(* IEC 61131-3 sources: brOscatLib/oscatBasic (part 4) *)

(* ---- FADE.st ---- *)
FUNCTION_BLOCK FADE
    (*http://www.oscat.de/images/OSCATBasic/oscat_basic333_en.pdf#page=276*)
    rmx(RST := RST AND NOT F, SET := RST AND F, PT := TF, UP := F);
    Y := (IN2 - IN1) / 65535.0 * WORD_TO_REAL(rmx.OUT) + IN1;

    (* code for rev 1.1
    IF RST THEN
    	rmx(set := F, RST := NOT F);
    ELSIF F AND (NOT rmx.high) THEN
    	rmx(PT := TF, UP := TRUE, e := TRUE, RST := FALSE, set := FALSE);
    ELSIF (NOT F) AND (NOT rmx.low) THEN
    	rmx(PT := TF, UP := FALSE, e := TRUE, RST := FALSE, set := FALSE);
    ELSE
    	rmx(e := FALSE, RST := FALSE, set := FALSE);
    END_IF
    Y := (WORD_TO_REAL(rmx.out) * IN1 + WORD_TO_REAL(FF - rmx.out) * IN2) / FF;
    *)

    (* revision history
    hm	26. dec 2007	rev 1.0
    	original version

    hm	18. oct. 2008	rev 1.1
    	improved performance
    	changed calls for rmp_w because rmp_w has chaged

    hm	17. dec. 2008	rev 1.2
    	function of input F was inverted

    hm	24. jan. 2009	rev 1.3
    	delted unused var FF
    *)
END_FUNCTION_BLOCK

(* ---- FF_D2E.st ---- *)
FUNCTION_BLOCK FF_D2E
    (*http://www.oscat.de/images/OSCATBasic/oscat_basic333_en.pdf#page=238*)
    IF RST THEN
    	Q0 := FALSE;
    	Q1 := FALSE;
    ELSIF CLK AND NOT edge_ THEN
    	Q0 := D0;
    	Q1 := D1;
    END_IF
    edge_ := CLK;

    (* revision history
    hm	25. dec 2007	rev 1.0
    	original version

    hm	27. dec 2007	rev 1.1
    	changed code for better performance

    hm	30. oct. 200	rev 1.2
    	deleted unnecessary init with 0

    hm	14. mar. 2009	rev 1.3
    	removed double assignments

    *)

END_FUNCTION_BLOCK

(* ---- FF_D4E.st ---- *)
FUNCTION_BLOCK FF_D4E
    (*http://www.oscat.de/images/OSCATBasic/oscat_basic333_en.pdf#page=239*)
    IF RST THEN
    	Q0 := FALSE;
    	Q1 := FALSE;
    	Q2 := FALSE;
    	Q3 := FALSE;
    ELSIF CLK AND NOT edge_ THEN
    	Q0 := D0;
    	Q1 := D1;
    	Q2 := D2;
    	Q3 := D3;
    END_IF
    edge_ := CLK;

    (* revision history
    hm	4. aug 2006	rev 1.0
    	original version

    hm	27. dec 2007	rev 1.1
    	changed code for better performance

    hm	30. oct. 200	rev 1.2
    	deleted unnecessary init with 0

    hm	14. mar. 2009	rev 1.3
    	removed double assignments

    *)

END_FUNCTION_BLOCK

(* ---- FF_DRE.st ---- *)
FUNCTION_BLOCK FF_DRE
    (*http://www.oscat.de/images/OSCATBasic/oscat_basic333_en.pdf#page=240*)
    IF RST OR SET THEN
    	Q := NOT RST;
    ELSIF CLK AND NOT edge_ THEN
    	Q := D;
    END_IF
    edge_ := CLK;

    (* revision history
    hm	4. aug 2006		rev 1.0
    	original version

    hm	27. dec 2007	rev 1.1
    	changed code for better performance

    hm	30. oct. 2008	rev 1.2
    	optimized performance
    *)
END_FUNCTION_BLOCK

(* ---- FF_JKE.st ---- *)
FUNCTION_BLOCK FF_JKE
    (*http://www.oscat.de/images/OSCATBasic/oscat_basic333_en.pdf#page=241*)
    IF RST OR SET THEN
    	Q := NOT RST;
    ELSIF CLK AND NOT edge_ THEN
    	IF J XOR K THEN Q := J;
    	ELSE Q := K XOR Q;
    	END_IF
    END_IF
    edge_ := CLK;

    (* revision history
    hm	4. aug 2006		rev 1.0
    	original version

    hm	27. dec 2007	rev 1.1
    	changed code for better performance

    hm	30. oct. 2008	rev 1.2
    	optimized performance
    *)
END_FUNCTION_BLOCK

(* ---- FF_RSE.st ---- *)
FUNCTION_BLOCK FF_RSE
    (*http://www.oscat.de/images/OSCATBasic/oscat_basic333_en.pdf#page=242*)
    IF RST THEN
    	(* asynchronous reset *)
    	Q := FALSE;
    ELSIF CR AND NOT er THEN
    	(* rising edge on CR *)
    	Q := FALSE;
    ELSIF CS AND NOT es THEN
    	(* rising edge on CS *)
    	Q := TRUE;
    END_IF

    es := CS;
    er := CR;

    (* revision history

    hm	16. jul. 2008	rev 1.0
    	original version

    *)

END_FUNCTION_BLOCK

(* ---- FIFO_16.st ---- *)
FUNCTION_BLOCK FIFO_16
    (*http://www.oscat.de/images/OSCATBasic/oscat_basic333_en.pdf#page=184*)
    IF RST THEN
    	pw := pr;
    	FULL := FALSE;
    	EMPTY := TRUE;
    	DOUT := 0;
    ELSIF E THEN
    	IF NOT EMPTY AND RD THEN
    		DOUT := fifo[pr];
    		pr := INC1(pr,n);
    		EMPTY := pr = pw;
    		FULL := FALSE;
    	END_IF
    	IF NOT FULL AND WD THEN
    		fifo[pw] := DIN;
    		pw := INC1(pw,n);
    		FULL := pw = pr;
    		EMPTY := FALSE;
    	END_IF
    END_IF

    (* revision history

    hm	4. aug. 2006	rev 1.0
    	original version

    hm	19. feb 2008	rev 1.1
    	performance improvements

    hm	17. oct. 2008	rev 1.2
    	improved performance

    ks	27. oct. 2008	rev 1.3
    	optimized coding

    hm	14. mar. 2009	rev 1.4
    	removed double assignments

    hm 24. jul. 2009	rev 2.0
    	chaged inputs E and WR to E, WD and WR
    	allow read and write in one cycle

    *)

END_FUNCTION_BLOCK

(* ---- FIFO_32.st ---- *)
FUNCTION_BLOCK FIFO_32
    (*http://www.oscat.de/images/OSCATBasic/oscat_basic333_en.pdf#page=184*)
    IF RST THEN
    	pw := pr;
    	FULL := FALSE;
    	EMPTY := TRUE;
    	DOUT := 0;
    ELSIF E THEN
    	IF NOT EMPTY AND RD THEN
    		DOUT := fifo[pr];
    		pr := INC1(pr,n);
    		EMPTY := pr = pw;
    		FULL := FALSE;
    	END_IF
    	IF NOT FULL AND WD THEN
    		fifo[pw] := DIN;
    		pw := INC1(pw,n);
    		FULL := pw = pr;
    		EMPTY := FALSE;
    	END_IF
    END_IF

    (* revision history
    hm	4. aug. 2006	rev 1.0
    	original version

    hm	19. feb 2008	rev 1.1
    	performance improvements

    hm	17. oct. 2008	rev 1.2
    	improved performance

    ks	27. oct. 2008 rev 1.3
    	improved code

    hm	14. mar. 2009	rev 1.4
    	removed double assignments

    hm 24. jul. 2009	rev 2.0
    	chaged inputs E and WR to E, WD and WR
    	allow read and write in one cycle

    *)

END_FUNCTION_BLOCK

(* ---- FILTER_DW.st ---- *)
FUNCTION_BLOCK FILTER_DW
    (*http://www.oscat.de/images/OSCATBasic/oscat_basic333_en.pdf#page=277*)
    (* read system time *)
    tx := T_PLC_MS();

    (* startup initialisation *)
    IF NOT init OR T = T#0s THEN
    	init := TRUE;
    	Yi := UDINT_TO_REAL(X);
    ELSE
    	Yi := Yi + (UDINT_TO_REAL(X) - UDINT_TO_REAL(Y)) * UDINT_TO_REAL(tx - last) / TIME_TO_REAL(T);
    END_IF
    last := tx;

    Y := REAL_TO_UDINT(Yi);

    (*
    hm 10. oct. 2008	rev 1.0
    	original version

    hm	3. nov. 2008	REV 1.1
    	corrected an overflow problem
    *)
END_FUNCTION_BLOCK

(* ---- FILTER_I.st ---- *)
FUNCTION_BLOCK FILTER_I
    (*http://www.oscat.de/images/OSCATBasic/oscat_basic333_en.pdf#page=278*)
    (* read system time *)
    tx := T_PLC_MS();

    (* startup initialisation *)
    IF NOT init OR T = T#0s THEN
    	init := TRUE;
    	Yi := INT_TO_DINT(X) * 1000;
    ELSE
    	(* to increase accuracy of the filter we calculate internal Yi wich is Y * 1000 *)
    	Yi := Yi + INT_TO_DINT(X - Y) * UDINT_TO_DINT(tx - last) * 1000 / TIME_TO_DINT(T);
    END_IF
    last := tx;
    Y := DINT_TO_INT(Yi / 1000);

    (*
    hm 8. nov. 2008	rev 1.0
    	original version

    *)
END_FUNCTION_BLOCK

(* ---- FILTER_MAV_DW.st ---- *)
FUNCTION_BLOCK FILTER_MAV_DW
    (*http://www.oscat.de/images/OSCATBasic/oscat_basic333_en.pdf#page=278*)
    (* limit N to size of buffer *)
    N := MIN(N, 32);

    (* startup initialisation *)
    IF NOT init OR RST OR N = 0 THEN
    	init := TRUE;
    	tmp := UINT_TO_INT(N)-1;
    	FOR i := 0 TO tmp DO
    		buffer[i] := DWORD_TO_UDINT(X);
    	END_FOR
    	Y := X;
    ELSE
    	tmp := UINT_TO_INT(N);
    	i := INC1(i, tmp);
    	Y := UDINT_TO_DWORD(DWORD_TO_UDINT(Y) + (DWORD_TO_UDINT(X) - buffer[i]) / N);
    	buffer[i] := DWORD_TO_UDINT(X);
    END_IF

    (*
    hm 13. oct. 2008	rev 1.0
    	original version

    hm	27. oct. 2008	rev 1.1
    	added typecast to avoid warnings

    hm	24. nov. 2008	rev 1.2
    	added typecasts to avoid warnings
    	avoid divide by 0 if N = 0

    hm	23. feb. 2009	rev 1.3
    	limit N to max array size

    *)
END_FUNCTION_BLOCK

(* ---- FILTER_MAV_W.st ---- *)
FUNCTION_BLOCK FILTER_MAV_W
    (*http://www.oscat.de/images/OSCATBasic/oscat_basic333_en.pdf#page=279*)
    (* limit N to size of buffer *)
    N := MIN(N, 32);

    (* startup initialisation *)
    IF NOT init OR RST OR N = 0 THEN
    	init := TRUE;
    	tmp := UINT_TO_INT(N) - 1;
    	FOR i := 1 TO tmp DO
    		buffer[i] := WORD_TO_UINT(X);
    	END_FOR
    	sum := WORD_TO_UINT(Y) * N;
    	Y := X;
    ELSE
    	tmp := UINT_TO_INT(N);
    	i := INC1(i, tmp);
    	sum := sum + WORD_TO_UINT(X) - buffer[i];
    	Y := UDINT_TO_WORD(sum / N);
    	buffer[i] := WORD_TO_UINT(X);
    END_IF

    (*
    hm 13. oct. 2008	rev 1.0
    	original version

    hm	18. oct. 2008	rev 1.1
    	added typecast to avoid warnings

    hm	24. nov. 2008	rev 1.2
    	added typecasts to avoid warnings
    	avoid devide by 0 if N = 0

    hm	23. feb. 2009	rev 1.3
    	limit N to max array size

    hm	26. mar. 2011	rev 1.4
    	corrected error in calculation
    *)
END_FUNCTION_BLOCK

(* ---- FILTER_W.st ---- *)
FUNCTION_BLOCK FILTER_W
    (*http://www.oscat.de/images/OSCATBasic/oscat_basic333_en.pdf#page=280*)
    (* read system time *)
    tx := T_PLC_MS();

    (* startup initialisation *)
    IF NOT init OR T = T#0s THEN
    	init := TRUE;
    	last := tx;
    	Y := X;
    ELSIF Y = X THEN
    	last := tx;
    ELSE
    	tmp :=  (WORD_TO_UINT(X) - WORD_TO_UINT(Y)) * (tx - last) / TIME_TO_UDINT(T);
    	IF tmp <> 0 THEN
    		Y := DINT_TO_WORD(WORD_TO_DINT(Y) + UDINT_TO_DINT(tmp));
    		last := tx;
    	END_IF
    END_IF

    (*
    hm 10. oct. 2008	rev 1.0
    	original version

    hm	3. nov. 2008	rev 1.1
    	fixed overflow problem in formula

    hm	25. jan. 2011	rev 1.2
    	fixed error in formula
    *)
END_FUNCTION_BLOCK

(* ---- FILTER_WAV.st ---- *)
FUNCTION_BLOCK FILTER_WAV
    (*http://www.oscat.de/images/OSCATBasic/oscat_basic333_en.pdf#page=280*)
    (* startup initialisation *)
    IF NOT init OR RST THEN
    	init := TRUE;
    	FOR i := 0 TO 15 DO
    		buffer[i] := X;
    	END_FOR
    	i := 15;
    	Y := X;
    ELSE
    	i := INC1(i, 16);
    	buffer[i] := X;
    END_IF

    (* calculate the weighted average *)
    Y := 0.0;
    FOR n := 0 TO 15 DO
    	Y := buffer[i] * W[n] + Y;
    	i := DEC1(i, 16);
    END_FOR

    (*
    hm 	14. oct. 2008	rev 1.0
    	original version

    hm	27. oct. 2008	rev 1.1
    	changed _DEC and _INC to DEC1 and INC1

    hm	10. mar. 2009	rev 1.2
    	real constants updated to new systax using dot

    *)

END_FUNCTION_BLOCK

(* ---- FLOW_CONTROL.st ---- *)
FUNCTION_BLOCK FLOW_CONTROL
    (*http://www.oscat.de/images/OSCATBasic/oscat_basic333_en.pdf#page=456*)
    STATUS := 100;
    IF RST THEN
    	Q := FALSE;
    	timer(RST := TRUE);
    	timer.RST := FALSE;
    	STATUS := 103;
    ELSIF ENQ THEN
    	IF IN THEN
    		STATUS := 101;
    	END_IF
    	IF REQ THEN
    		(* timer will generate a timed pulse after TP goes high *)
    		timer.PT1 := T_AUTO;
    		timer.PTD := T_DELAY;
    		timer.IN := TRUE;
    		STATUS := 102;
    	END_IF
    END_IF

    (* set output and run timer *)
    timer();
    timer.IN := FALSE;
    Q := (IN AND ENQ) OR timer.Q;

    (* revision history
    hm 	28. jun. 2008 	rev 1.0
    	original version

    *)
END_FUNCTION_BLOCK

(* ---- FLOW_METER.st ---- *)
FUNCTION_BLOCK FLOW_METER
    (*http://www.oscat.de/images/OSCATBasic/oscat_basic333_en.pdf#page=339*)
    IF NOT init THEN	(* init on power up *)
    	init := TRUE;
    	tl := tx;
    	x_last := X;
    	y_last := Y;
    	int1.K := 2.7777777777777777E-4;
    END_IF

    (* run integrator *)
    int1(E := NOT (RST OR PULSE_MODE) AND E, X := VX, Y := X);	(* gated operation *)

    IF RST THEN		(* reset *)
    	X := 0.0;
    	Y := 0;
    	tl := tx;
    	x_last := 0.0;
    	y_last := 0;
    ELSIF E AND PULSE_MODE THEN	(* check for pulse mode *)
    	IF NOT e_last THEN X := X + VX; END_IF
    END_IF
    e_last := E;

    (* reduce X to be less than 1 and increase Y respectively *)
    IF X > 1.0 THEN
    	tmp := FLOOR(X);
    	Y := Y + INT_TO_UDINT(tmp);
    	X := X - INT_TO_REAL(tmp);
    END_IF

    (* calculate the current flow *)
    tx := UDINT_TO_TIME(T_PLC_MS());
    IF tx - tl >= UPDATE_TIME AND UPDATE_TIME > t#0s THEN
    	F := (UDINT_TO_REAL(Y - y_last) + X - x_last) / TIME_TO_REAL(tx - tl) * 3.6E6;
    	y_last := Y;
    	x_last := X;
    	tl := tx;
    END_IF

    (* revision history
    hm	23. jan. 2011	rev 1.0
    	original version

    *)

END_FUNCTION_BLOCK

(* ---- FT_AVG.st ---- *)
FUNCTION_BLOCK FT_AVG
    (*http://www.oscat.de/images/OSCATBasic/oscat_basic333_en.pdf#page=98*)
    (* limit N to a max of 32 because delay can do max 32 cycles *)
    buff.N := LIMIT(0, N, 32);

    IF NOT init OR RST THEN
    	FOR i := 1 TO N DO
    		buff(IN := IN);
    	END_FOR
    	AVG := IN;
    	init := TRUE;
    ELSIF E THEN
    	buff(IN := IN);
    	AVG := AVG + (IN - buff.OUT ) / INT_TO_REAL(N);
    END_IF

    (* revision history

    hm	7. jan. 2007	rev 1.1
    	chaged RST logic to load the buffer with the actual input value instead of 0.
    	added en input to allow better control of signal flow
    	added init to load the buffer with IN at startup to avoid rampup at beginning.
    	deleted unused variable cnt.

    hm	14. jun. 2008	rev 1.2
    	set default for input en = TRUE and N = 32

    hm	10. oct. 2008	rev 1.3
    	improved performance

    hm	18. oct. 2008	rev 1.4
    	changed input en to E for compatibility reasons

    hm	10. mar. 2009	rev 1.5
    	added type conversion for compatibility reasons

    *)
END_FUNCTION_BLOCK

(* ---- FT_DERIV.st ---- *)
FUNCTION_BLOCK FT_DERIV
    (*http://www.oscat.de/images/OSCATBasic/oscat_basic333_en.pdf#page=396*)
    (* read system time *)
    tx := T_PLC_US();
    tc := UDINT_TO_REAL(tx - last);
    last := tx;

    (* init on first startup *)
    IF NOT init THEN
    	init := TRUE;
    	old := IN;
    ELSIF RUN AND tc > 0.0 THEN
    	OUT := (IN - old) / tc * 1000000.0 * K;
    	old := IN;
    ELSE
    	OUT := 0.0;
    END_IF

    (*
    hm 3.1.2007			rev 1.1
    	added init code for startup
    	set the default for K to 1

    hm	15. sep 2007	rev 1.2
    	replaced Time() with T_PLC_US for compatibility and performance reasons
    	increased accuracy and work IN microseconds internally

    hm 29 oct 2007	rev 1.3
    	prohibit calculation when tx - last = 0 to avoid division by 0 and increase accuracy on fast systems

    hm	6. nov. 2008	rev 1.4
    	improved performance

    hm	11. mar. 2009	rev 1.5
    	inproved code
    *)
END_FUNCTION_BLOCK

(* ---- FT_IMP.st ---- *)
FUNCTION_BLOCK FT_IMP
    (*http://www.oscat.de/images/OSCATBasic/oscat_basic333_en.pdf#page=399*)
    t1(IN:= IN, T:=T);
    OUT := (IN - t1.OUT) * K;

    (*
    hm 3.1.2007	rev 1.1
    	added factor K

    *)
END_FUNCTION_BLOCK

(* ---- FT_INT.st ---- *)
FUNCTION_BLOCK FT_INT
    (*http://www.oscat.de/images/OSCATBasic/oscat_basic333_en.pdf#page=400*)
    IF RST THEN
    	OUT := 0.0;
    ELSE
    	INTeg(X := IN, E := RUN, K := K, Y := OUT);
    END_IF

    (* limit the outputs *)
    IF OUT >= OUT_MAX THEN
    	OUT := OUT_MAX;
    	LIM := TRUE;
    ELSIF OUT <= OUT_MIN THEN
    	OUT := OUT_MIN;
    	LIM := TRUE;
    ELSE
    	LIM := FALSE;
    END_IF

    (*
    hm 13.12.2006	rev 1.1
    	changed to "trapezregel" which increases accuracy
    	before OUT := OUT + IN * time new: OUT := OUT + (IN + in_last) / 2 * time

    hm 15.1.2007		rev 1.2
    	added default for K to be 1.

    hm	15.9.2007		rev 1.3
    	replaced time() with T_PLC_US for compatibility and performance reason
    	increased internal accuracy to microseconds

    hm 29. oct 2007		rev 1.4
    	changed code so int will not be called is time difference is 0 to increase accuracy on systems
    	with cycle times below 1ms

    hm	2. dec 2007	 	rev 1.5
    	changed code for better performance

    hm	5. jan 2008		rev 1.6
    	further improvements IN performance

    hm	8. feb 2008		rev 1.7
    	deleted limits +/- 1000 now limit is the range of real
    	added variables out1 and out2 to extend the resolution
    	corrected an error with elapsed time
    	deleted unusfull output ET

    hm	13. mar 2008	rev 1.8
    	changed preset value OUT_MIN to -1e37.
    	stop integrator at the limits.

    hm	16. mar 2008	rev 1.9
    	added type conversion to avoid warning under codesys 3.0

    hm	2. jun. 2008	rev 2.0
    	rewritten with clear code
    	limits can now be set without RUN

    hm	3. nov. 2008	rev 2.1
    	optimized code using INTEGRATE and LIMX

    hm	10. mar. 2009	rev 2.2
    	removed nested comments
    *)

END_FUNCTION_BLOCK

(* ---- FT_INT2.st ---- *)
FUNCTION_BLOCK FT_INT2
    (*http://www.oscat.de/images/OSCATBasic/oscat_basic333_en.pdf#page=402*)
    IF RST THEN
    	R2_SET(0.0, val);
    	OUT := 0.0;
    ELSE
    	integ(X := IN, E := RUN, K := K, Y := ix);
    	R2_ADD(val, ix, val);
    	ix := 0.0;
    	OUT := val.RX;
    END_IF

    (* check output for limits *)
    IF OUT > OUT_MIN AND OUT < OUT_MAX THEN
    	LIM := FALSE;
    ELSE
    	OUT := LIMIT(OUT_MIN, OUT, OUT_MAX);
    	R2_SET(OUT, val);
    	LIM := TRUE;
    END_IF

    (*	revision history
    hm	2. jun. 2008	rev 1.0
    	original version

    hm	5. nov. 2008	rev 1.1
    	rewritten code using integrate

    hm	11. mar. 2009	rev 1.2
    	real constants updated to new systax using dot

    *)

END_FUNCTION_BLOCK

(* ---- FT_MIN_MAX.st ---- *)
FUNCTION_BLOCK FT_MIN_MAX
    (*http://www.oscat.de/images/OSCATBasic/oscat_basic333_en.pdf#page=99*)
    IF RST OR NOT init THEN
    	MN := IN;
    	MX := IN;
    	init := TRUE;
    ELSIF IN < MN THEN MN := IN;
    ELSIF IN > MX THEN MX := IN;
    END_IF
END_FUNCTION_BLOCK

(* ---- FT_PD.st ---- *)
FUNCTION_BLOCK FT_PD
    (*http://www.oscat.de/images/OSCATBasic/oscat_basic333_en.pdf#page=403*)
    (* run differentiator *)
    diff(IN := IN, K := TV);

    (* combine both values *)
    Y := KP * (diff.OUT + IN);

    (* revision history
    hm 	3. jun. 2008 	rev 1.0
    	original version

    *)
END_FUNCTION_BLOCK

(* ---- FT_PDT1.st ---- *)
FUNCTION_BLOCK FT_PDT1
    (*http://www.oscat.de/images/OSCATBasic/oscat_basic333_en.pdf#page=403*)
    (* run differentiator *)
    diff(IN := IN, K := TV);

    (* Run PT1 filter *)
    TP(IN := diff.OUT, T := REAL_TO_TIME(T1));

    (* combine both values *)
    Y := KP * (TP.OUT + IN);

    (* revision history
    hm 	3. jun. 2008 	rev 1.0
    	original version

    *)
END_FUNCTION_BLOCK

(* ---- FT_PI.st ---- *)
FUNCTION_BLOCK FT_PI
    (*http://www.oscat.de/images/OSCATBasic/oscat_basic333_en.pdf#page=404*)
    (* run integrator *)
    integ(IN := IN, K := KI, RUN := IEN, RST := RST, OUT_MIN := ILIM_L, OUT_MAX := ILIM_H);

    (* check if integrator has reached its limits and set overflow *)
    LIM := integ.LIM;
    Y := KP * IN + integ.OUT;

    (* revision history
    hm 	3. jun. 2008 	rev 2.0
    	original version

    *)
END_FUNCTION_BLOCK

(* ---- FT_PID.st ---- *)
FUNCTION_BLOCK FT_PID
    (*http://www.oscat.de/images/OSCATBasic/oscat_basic333_en.pdf#page=406*)
    (* run integrator only if TN > 0 *)
    IF TN > 0.0 THEN
    	integ(IN := IN, K := 1.0 / TN, RUN := IEN, RST := RST, OUT_MIN := ILIM_L, OUT_MAX := ILIM_H);
    ELSE
    	integ(RST := FALSE);
    END_IF

    (* run differentiator *)
    diff(IN := IN, K := TV);

    (* combine both values *)
    Y := KP * (integ.OUT + diff.OUT + IN);

    (* check if integrator has reached its limits and set overflow *)
    LIM := integ.LIM;

    (* revision history
    hm 3. jun. 2008 	rev 2.0
    	original version

    hm	11. mar. 2009	rev 2.1
    	real constants updated to new systax using dot

    *)
END_FUNCTION_BLOCK

(* ---- FT_PIDW.st ---- *)
FUNCTION_BLOCK FT_PIDW
    (*http://www.oscat.de/images/OSCATBasic/oscat_basic333_en.pdf#page=407*)
    (* run the integrator *)
    IF TN = 0.0 OR RST THEN
    	integ(E := FALSE, Y := YI);
    	YI := 0.0;
    ELSE
    	integ(X := IN, K := 1.0 / TN, E := NOT LIM, Y := YI);
    END_IF

    (* add up integrator and linear part *)
    Y := KP * (IN + YI);

    (* run differentiator *)
    diff(IN := IN, K := TV);

    (* set LIM before differentiator is added to stop integrator if necessary *)
    IF Y > LIM_L AND Y < LIM_H THEN
    	LIM := FALSE;
    ELSE
    	LIM := TRUE;
    END_IF

    (* add differential part and limit output Y *)

    Y := LIMIT(LIM_L, Y + KP * diff.OUT, LIM_H);

    (* revision history
    hm 3. jun. 2008 	rev 1.0
    	original version

    hm	5. nov. 2008	rev 1.1
    	changed code to use integrate

    hm	11. mar. 2009	rev 1.2
    	real constants updated to new systax using dot

    *)
END_FUNCTION_BLOCK

(* ---- FT_PIDWL.st ---- *)
FUNCTION_BLOCK FT_PIDWL
    (*http://www.oscat.de/images/OSCATBasic/oscat_basic333_en.pdf#page=409*)
    (* if RST then *)
    IF RST THEN
    	piwl(RST := TRUE);
    	piwl.RST := FALSE;
    ELSE
    	(* run piwl controller first *)
    	(* we need to check if TN = 0 and do alternative calls *)
    	IF TN = 0.0 THEN
    		piwl(IN := IN * KP, KP := 1.0, KI := 0.0, LIM_L := LIM_L, LIM_H := LIM_H);
    	ELSE
    		piwl(IN := IN * KP, KP := 1.0, KI := 1.0 / TN, LIM_L := LIM_L, LIM_H := LIM_H);
    	END_IF

    	(* run differentiator and add_to_output *)
    	diff(IN := IN, K := KP * TV);
    	Y := piwl.Y + diff.OUT;

    	(* limit the output *)
    	IF Y < LIM_L THEN
    		LIM := TRUE;
    		Y := LIM_L;
    	ELSIF Y > LIM_H THEN
    		LIM := TRUE;
    		Y := LIM_H;
    	ELSE
    		LIM := FALSE;
    	END_IF
    END_IF

    (* revision history
    hm 13. jun. 2008 	rev 1.0
    	original version

    hm	25. jan 2008	rev 1.1
    	multiply differential part with KP

    hm	11. mar. 2009	rev 1.2
    	real constants updated to new systax using dot

    hm	13. nov. 2009	rev 1.3
    	fixed code for negative KP

    *)
END_FUNCTION_BLOCK

(* ---- FT_PIW.st ---- *)
FUNCTION_BLOCK FT_PIW
    (*http://www.oscat.de/images/OSCATBasic/oscat_basic333_en.pdf#page=411*)
    (* run integrator *)
    integ(IN := IN, K := KI, RUN := NOT LIM, RST := RST);

    (* set output value *)
    Y := KP * IN + integ.OUT;

    (* check for limits and set integrator for anti wind up *)
    IF Y < LIM_L THEN
    	Y := LIM_L;
    	LIM := TRUE;
    ELSIF Y > LIM_H THEN
    	Y := LIM_H;
    	LIM := TRUE;
    ELSE
    	LIM := FALSE;
    END_IF

    (* revision history
    hm 	3. jun. 2008 	rev 1.0
    	original version

    *)
END_FUNCTION_BLOCK

(* ---- FT_PIWL.st ---- *)
FUNCTION_BLOCK FT_PIWL
    (*http://www.oscat.de/images/OSCATBasic/oscat_basic333_en.pdf#page=412*)
    (* initialize at power_up *)
    IF NOT init OR RST THEN
    	init := TRUE;
    	in_last := IN;
    	t_last := T_PLC_US();
    	i := 0.0;
    	tc := 0.0;
    ELSE
    	(* read last cycle time IN Microseconds *)
    	tx := T_PLC_US();
    	tc := UDINT_TO_REAL(tx - t_last);
    	t_last := tx;

    	(* calculate proportional part *)
    	p := KP * IN;

    	(* run integrator *)
    	i := (IN + in_last) * 5.0E-7 * KI * tc + i;
    	in_last := IN;

    	(* calculate output Y *)
    	Y := p + i;

    	(* check output for limits *)
    	IF Y >= LIM_H THEN
    		Y := LIM_H;
    		IF KI <> 0.0 THEN
    			i := LIM_H - p;
    		ELSE
    			i := 0.0;
    		END_IF
    		LIM := TRUE;
    	ELSIF Y <= LIM_L THEN
    		Y := LIM_L;
    		IF KI <> 0.0 THEN
    			i := LIM_L - p;
    		ELSE
    			i := 0.0;
    		END_IF
    		LIM := TRUE;
    	ELSE
    		LIM := FALSE;
    	END_IF
    END_IF

    (* revision history
    hm 13. jun. 2008 	rev 1.0
    	original version

    hm	27. oct. 2008	rev 1.1
    	integrator will not be adjusted when KI = 0

    hm	25. jan 2009	rev 1.2
    	module will also work with negative K

    hm	11. mar. 2009	rev 1.3
    	real constants updated to new systax using dot

    *)
END_FUNCTION_BLOCK

(* ---- FT_Profile.st ---- *)
FUNCTION_BLOCK FT_Profile
    (*http://www.oscat.de/images/OSCATBasic/oscat_basic333_en.pdf#page=457*)
    (* read system time *)
    tx := UDINT_TO_TIME(T_PLC_MS());

    (* determine start condition *)
    IF E AND NOT edge_ THEN
    	RUN := TRUE;
    	ET := t#0s;
    	t0 := tx;
    	ta := tx;
    	tb := MULTIME(TIME_1, M);
    	va := VALUE_0;
    	vb := VALUE_1;
    	temp := VALUE_0;
    	state := 1;
    END_IF
    edge_ := E;

    (* generate startup profile *)
    IF RUN THEN
    	CASE state OF
    		1:	IF tx - ta >= tb THEN
    				ta := ta + tb;
    				tb := MULTIME(TIME_2 - TIME_1, M);
    				va := VALUE_1;
    				vb := VALUE_2;
    				temp := VALUE_1;
    				state := 2;
    			ELSE
    				temp := ((vb - va) * TIME_TO_REAL(tx - ta) / TIME_TO_REAL(tb) + va);
    			END_IF
    		2:	IF tx - ta >= tb THEN
    				ta := ta + tb;
    				tb := MULTIME(TIME_3 - TIME_2, M);
    				va := VALUE_2;
    				vb := VALUE_3;
    				temp := VALUE_2;
    				state := 3;
    			ELSE
    				temp := ((vb - va) * TIME_TO_REAL(tx - ta) / TIME_TO_REAL(tb) + va);
    			END_IF
    		3:	IF tx - ta >= tb THEN
    				ta := ta + tb;
    				tb := MULTIME(TIME_10 - TIME_3, M);
    				va := VALUE_3;
    				vb := VALUE_10;
    				temp := VALUE_3;
    				state := 4;
    			ELSE
    				temp := ((vb - va) * TIME_TO_REAL(tx - ta) / TIME_TO_REAL(tb) + va);
    			END_IF
    		4 :	IF tx - ta >= tb THEN
    				ta := ta + tb;
    				tb := MULTIME(TIME_11 - TIME_10, M);
    				va := VALUE_10;
    				vb := VALUE_11;
    				temp := VALUE_10;
    				IF E THEN state := 5; ELSE state := 6; END_IF
    			ELSE
    				temp := ((vb - va) * TIME_TO_REAL(tx - ta) / TIME_TO_REAL(tb) + va);
    			END_IF
    		5:	(* extend the signal while E is true *)
    			IF E THEN
    				ta := tx;
    			ELSE
    				state := 6;
    			END_IF
    		6:	IF tx - ta >= tb THEN
    				ta := ta + tb;
    				tb := MULTIME(TIME_12 - TIME_11, M);
    				va := VALUE_11;
    				vb := VALUE_12;
    				temp := VALUE_11;
    				state := 7;
    			ELSE
    				temp := ((vb - va) * TIME_TO_REAL(tx - ta) / TIME_TO_REAL(tb) + va);
    			END_IF
    		7:	IF tx - ta >= tb THEN
    				ta := ta + tb;
    				tb := MULTIME(TIME_13 - TIME_12, M);
    				va := VALUE_12;
    				vb := VALUE_13;
    				temp := VALUE_12;
    				state := 8;
    			ELSE
    				temp := ((vb - va) * TIME_TO_REAL(tx - ta) / TIME_TO_REAL(tb) + va);
    			END_IF
    		8:	IF tx - ta >= tb THEN
    				temp := VALUE_13;
    				RUN := FALSE;
    			ELSE
    				temp := ((vb - va) * TIME_TO_REAL(tx - ta) / TIME_TO_REAL(tb) + va);
    			END_IF
    	END_CASE
    	Y := temp * K + O;
    	ET := tx - t0;
    END_IF

    (* revision history
    hm	27 feb 2007		rev 1.0
    	original version

    hm	15. sep2007		rev 1.1
    	replaced Time() with T_PLC_MS for compatibility and performance reasons

    *)
END_FUNCTION_BLOCK

(* ---- FT_PT1.st ---- *)
FUNCTION_BLOCK FT_PT1
    (*http://www.oscat.de/images/OSCATBasic/oscat_basic333_en.pdf#page=414*)
    (* read system time *)
    tx := T_PLC_US();

    (* startup initialisation *)
    IF NOT init OR T = T#0s THEN
    	init := TRUE;
    	OUT := K * IN;
    ELSE
    	OUT := OUT + (IN * K - OUT) * UDINT_TO_REAL(tx - last) / TIME_TO_REAL(T) * 1.0E-3;
    	IF ABS(OUT) < 1.0E-20 THEN OUT := 0.0; END_IF
    END_IF
    last := tx;

    (*
    hm 1.1.2007	rev 1.1
    	corrected error while startup value was not correct
    	for very small time values real output would run OUT of range.

    hm 3.1.2007	rev 1.2
    	corrected an error for falling edge failures.
    	added output faktor K.

    hm 27. 2. 2007	rev 1.3
    	output will be input during init for definitive startup condition.

    hm	15.9.2007	rev 1.4
    	changed time() to T_PLC_US() for compatibilitxy resons
    	increased internal accuracy to Microseconds instead of Milliseconds

    hm	23. oct 2007	rev 1.5
    	added OUT := IN to the init statements

    hm	30. nov 2007	rev 1.6
    	changed OUT to be K * IN during initialization

    hm	5. jan 2008	rev 1.7
    	improved code for better performance

    hm	16. mar. 2008	rev 1.8
    	added type conversion to avoid warning under codesys 3.0

    hm	14. jun. 2008	rev 1.9
    	improved code

    hm	11. mar. 2009	rev 1.10
    	real constants updated to new systax using dot

    hm	18. jan. 2011	rev 1.11
    	avoid underrun of OUT
    *)
END_FUNCTION_BLOCK

(* ---- FT_PT2.st ---- *)
FUNCTION_BLOCK FT_PT2
    (*http://www.oscat.de/images/OSCATBasic/oscat_basic333_en.pdf#page=415*)
    (* startup initialisation *)
    IF NOT init OR T = T#0s THEN
    	init := TRUE;
    	OUT := K * IN;
    	I2 := OUT;
    ELSE
    	tn := TIME_TO_REAL(T) * 1.0E-3;
    	tn2 := tn * tn;
    	int1(X := IN * K / tn2 - I1 * 0.5 * D / tn - I2 / tn2, Y := I1);
    	int2(X := I1,Y := I2);
    	OUT := I2;
    END_IF

    (* revision history

    15.1.2007 hm		rev 1.1
    	changed formula to new more acurate formula

    hm 15.9.2007		rev 1.2
    	deleted unused code for init system time reading tx

    hm	30.11.2007	rev 1.3
    	changed OUT to be K * IN during initialization
    	avoind divide by 0 if tn = 0

    hm	3. nov. 2008	rev 1.4
    	optimized code and fixed a problem with init

    hm	11. mar. 2009	rev 1.5
    	real constants updated to new systax using dot

    *)
END_FUNCTION_BLOCK

(* ---- FT_RMP.st ---- *)
FUNCTION_BLOCK FT_RMP
    (*http://www.oscat.de/images/OSCATBasic/oscat_basic333_en.pdf#page=100*)
    (* read system time *)
    tx := UDINT_TO_TIME(T_PLC_MS()) - last;

    IF NOT init THEN
    	init := TRUE;
    	last := tx;
    	tx := t#0s;
    	OUT := IN;
    END_IF
    IF NOT RMP THEN
    	OUT := IN;
    	BUSY := FALSE;
    ELSIF OUT > IN THEN
    	(* ramp down *)
    	OUT := OUT - TIME_TO_REAL(tx) * 0.001 * KF;
    	OUT := MAX(IN, OUT);
    ELSIF OUT < IN THEN
    	(* ramp up *)
    	OUT := OUT + TIME_TO_REAL(tx) * 0.001 * KR;
    	OUT := MIN(IN, OUT);
    END_IF

    (* set BUSY and dir flags *)
    IF OUT < IN THEN
    	BUSY := TRUE;
    	UD := TRUE;
    ELSIF OUT > IN THEN
    	BUSY := TRUE;
    	UD := FALSE;
    ELSE
    	BUSY := FALSE;
    END_IF
    last := last + tx;

    (* revision history:

    hm 8.10.2006			rev 1.1
    	added UD output

    hm 12. feb 2007		rev 1.2
    	added init variable and corrected a possible startup problem

    hm	17. sep 2007	rev 1.3
    	replaced time() with t_plc_ms() for compatibility reasons

    hm	25. jan 2008	rev 1.4
    	performance improvements
    	allow KR and KF to be 0
    *)
END_FUNCTION_BLOCK

(* ---- FT_TN16.st ---- *)
FUNCTION_BLOCK FT_TN16
    (*http://www.oscat.de/images/OSCATBasic/oscat_basic333_en.pdf#page=416*)
    (* read system time *)
    tx := UDINT_TO_TIME(T_PLC_MS());

    TRIG := FALSE;
    IF NOT init THEN
    	X[cnt] := IN;
    	init := TRUE;
    	last := tx;
    ELSIF tx - last >= T / length THEN
    	IF cnt = length - 1 THEN cnt := 0; ELSE cnt := cnt + 1; END_IF
    	OUT := X[cnt];
    	X[cnt] := IN;
    	last := tx;
    	TRIG := TRUE;
    END_IF

    (* revision history
    hm		1. jan 2007	rev 1.0
    	original version

    hm		16. sep 2007	rev 1.1
    	changes time() to T_plc_ms() for compatibility reasons

    *)
END_FUNCTION_BLOCK

(* ---- FT_TN64.st ---- *)
FUNCTION_BLOCK FT_TN64
    (*http://www.oscat.de/images/OSCATBasic/oscat_basic333_en.pdf#page=419*)
    (* read system time *)
    tx := UDINT_TO_TIME(T_PLC_MS());

    TRIG := FALSE;
    IF NOT init THEN
    	X[cnt] := IN;
    	init := TRUE;
    	last := tx;
    ELSIF tx - last >= T / length THEN
    	IF cnt = length - 1 THEN cnt := 0; ELSE cnt := cnt + 1; END_IF
    	OUT := X[cnt];
    	X[cnt] := IN;
    	last := tx;
    	TRIG := TRUE;
    END_IF

    (* revision history
    hm		1. jan 2007		rev 1.0
    	original version

    hm		16. sep 2007	rev 1.1
    	changes time() to T_plc_ms() for compatibility reasons

    *)
END_FUNCTION_BLOCK

(* ---- FT_TN8.st ---- *)
FUNCTION_BLOCK FT_TN8
    (*http://www.oscat.de/images/OSCATBasic/oscat_basic333_en.pdf#page=420*)
    tx := UDINT_TO_TIME(T_PLC_MS());
    TRIG := FALSE;
    IF NOT init THEN
    	X[cnt] := IN;
    	init := TRUE;
    	last := tx;
    ELSIF tx - last >= T / length THEN
    	IF cnt = length - 1 THEN cnt := 0; ELSE cnt := cnt + 1; END_IF
    	OUT := X[cnt];
    	X[cnt] := IN;
    	last := tx;
    	TRIG := TRUE;
    END_IF

    (* revision history
    hm		1. jan 2007		rev 1.0
    	original version

    hm		16. sep 2007	rev 1.1
    	changes time() to T_plc_ms() for compatibility reasons

    *)
END_FUNCTION_BLOCK

(* ---- GEN_BIT.st ---- *)
FUNCTION_BLOCK GEN_BIT
    (*http://www.oscat.de/images/OSCATBasic/oscat_basic333_en.pdf#page=196*)
    (* check if number of runs is finished or REP = 0 which means continuous *)

    IF CLK AND NOT RST THEN
    	RUN := (REP = 0) OR (rx <= REP);
    	IF RUN THEN
    		(* check for step counter reached and reset to 0 if CNT = STEPS *)
    		IF CNT = STEPS THEN
    			CNT := 0;
    		END_IF

    		(* when CNT = 0 then reload the inputs into the registers *)
    		IF CNT = 0 THEN
    			r0 := IN0;
    			r1 := IN1;
    			r2 := IN2;
    			r3 := IN3;
    		END_IF

    		(* when CNT < STEPS, shift the lowest bits to the outputs *)
    		IF (CNT < STEPS) THEN
    			Q0 := r0.0;
    			Q1 := r1.0;
    			Q2 := r2.0;
    			Q3 := r3.0;
    			r0 := SHR(r0,1);
    			r1 := SHR(r1,1);
    			r2 := SHR(r2,1);
    			r3 := SHR(r3,1);
    		END_IF

    		(* increment the step counter *)
    		CNT := CNT +1;
    		IF (CNT = STEPS) AND (REP <> 0) THEN rx := rx +1; END_IF
    		IF (rx > REP) AND (REP <> 0) THEN RUN := FALSE; END_IF
    	END_IF
    ELSE
    	IF RST THEN
    		RUN := FALSE;
    		Q0 := FALSE;
    		Q1 := FALSE;
    		Q2 := FALSE;
    		Q3 := FALSE;
    		r0 := 0;
    		r1 := 0;
    		r2 := 0;
    		r3 := 0;
    		CNT := 0;
    		rx := 1;
    	END_IF
    END_IF

    (* revision histroy
    hm	4 aug 2006	rev 1.0
    	original version

    hm 15. oct. 2008	rev 1.1
    	improved performance

    hm	14. mar. 2009	rev 1.2
    	removed double assignments

    *)
END_FUNCTION_BLOCK

(* ---- GEN_PULSE.st ---- *)
FUNCTION_BLOCK GEN_PULSE
    (*http://www.oscat.de/images/OSCATBasic/oscat_basic333_en.pdf#page=257*)
    IF ENQ THEN
    	tx := UDINT_TO_TIME(T_PLC_MS());
    	IF NOT init THEN init := TRUE; tn := tx; END_IF
    	IF tx - tn >= SEL(Q, PTL, PTH) THEN
    		tn := tn + SEL(Q, PTL, PTH);
    		Q := NOT Q;
    	END_IF
    ELSE
    	Q := FALSE;
    	init := FALSE;
    END_IF

    (* revision history
    hm	29. jun. 2008	rev 1.0
    	original version

    hm	23. nov. 2008	rev 1.1
    	set default for ENQ to be true

    hm	18. jul. 2009	rev 1.2
    	improved performance

    hm	13. nov. 2009	rev 1.3
    	corrected error

    hm	16. feb. 2011	rev 1.4
    	corrected an error when timer overflows

    hm	8. apr. 2011	rev 1.5
    	PTL and PTH was exchanged
    *)
END_FUNCTION_BLOCK

(* ---- GEN_PW2.st ---- *)
FUNCTION_BLOCK GEN_PW2
    (*http://www.oscat.de/images/OSCATBasic/oscat_basic333_en.pdf#page=258*)
    (* read system timer *)
    tx := UDINT_TO_TIME(T_PLC_MS());

    (* startup initialization *)
    IF NOT init THEN
    	start := tx;
    	init := TRUE;
    	TH := T#0s;
    	TL := T#0s;
    END_IF

    (* timing selection *)
    IF TS THEN
    	t_high := TH2;
    	t_low := TL2;
    ELSE
    	t_high := TH1;
    	t_low := TL1;
    END_IF

    (* normal operation *)
    IF ENQ THEN
    	et := tx - start;
    	IF NOT Q THEN
    		IF et >= t_low THEN
    			Q := TRUE;
    			start := tx;
    			TL := T#0s;
    		ELSE
    			TL := et;
    		END_IF
    	ELSE
    		IF et >= t_high THEN
    			Q := FALSE;
    			start := tx;
    			TH := T#0s;
    		ELSE
    			TH := et;
    		END_IF
    	END_IF
    ELSE
    	Q := FALSE;
    	TH := T#0s;
    	TL := T#0s;
    	start := tx;
    END_IF

    (* revision history
    hm	26. sep. 2008	rev 1.0
    	original version

    hm	14. mar. 2009	rev 1.1
    	removed double assignments

    *)
END_FUNCTION_BLOCK

(* ---- GEN_RDM.st ---- *)
FUNCTION_BLOCK GEN_RDM
    (*http://www.oscat.de/images/OSCATBasic/oscat_basic333_en.pdf#page=258*)
    (* read system time and prepare input data *)
    tx := UDINT_TO_TIME(T_PLC_MS()) - last;

    (* init section *)
    IF NOT init THEN
    	init := TRUE;
    	last := tx;
    	tx := t#0s;
    END_IF

    (* add last if one cycle is finished *)
    IF tx >= PT THEN
    	last := last + PT;
    	tx := tx - PT;

    	(* generate output signal *)
    	OUT := AM * (RDM(0) - 0.5) + OS;
    	Q := TRUE;
    ELSE
    	Q := FALSE;
    END_IF

    (* revision history

    hm	7.2.2007		rev 1.0
    	original version

    hm	16.9.2007		rev 1.1
    	changes time() to T_plc_ms() for compatibility reasons

    *)

END_FUNCTION_BLOCK

(* ---- GEN_RDT.st ---- *)
FUNCTION_BLOCK GEN_RDT
    (*http://www.oscat.de/images/OSCATBasic/oscat_basic333_en.pdf#page=259*)
    tonRDMTimer ( IN:= ENABLE , PT:= tRDMTime );
    tof_xQ ( IN:= tonRDMTimer.Q , PT:= TP_Q );
    XQ := tof_xQ.Q;
    IF tonRDMTimer.Q THEN
    		 XQ := TRUE ;
    		 rRDMTime := RDM (LAST:= rRDMTime ) ;
    		 tRDMTime := REAL_TO_TIME ( rRDMTime * DINT_TO_REAL(TIME_TO_DINT( MAX_TIME_MS - MIN_TIME_MS ) + TIME_TO_DINT(MIN_TIME_MS ))) ;
    		 tonRDMTimer ( IN:= FALSE );
    END_IF

    (* revision history
    J. Schohaus	19. nov 2007	rev 1.0
    	origial version

    hm	16. mar. 2008			rev 1.1
    	added type conversion to avoid warnings under codesys 3.0
    *)
END_FUNCTION_BLOCK

(* ---- GEN_RMP.st ---- *)
FUNCTION_BLOCK GEN_RMP
    (*http://www.oscat.de/images/OSCATBasic/oscat_basic333_en.pdf#page=260*)
    (* read system time and prepare input data *)
    tx := UDINT_TO_TIME(T_PLC_MS()) - last;
    DL := MODR(DL,1.0);
    IF DL < 0.0 THEN DL := 1.0 - DL; END_IF

    (* init section *)
    IF NOT init THEN
    	init := TRUE;
    	last := tx;
    	tx := t#0s;
    END_IF

    (* add last if one cycle is finished *)
    IF tx >= PT THEN
    	last := last + PT;
    	tx := tx - PT;
    END_IF

    (* generate sine wave *)
    ltemp := temp;
    IF PT > t#0s THEN temp := FRACT(TIME_TO_REAL(tx + MULTIME(PT, DL)) / TIME_TO_REAL(PT)); END_IF
    OUT := AM * temp + OS;

    (* boolean output Q *)
    Q := temp < ltemp;

    (* revision history
    hm	3. mar 2007		rev 1.0
    	original version

    hm	17 sep 2007		rev 1.1
    	replaced time() with t_plc_ms for compatibilitx reasons

    hm	27. nov 2007	rev 1.2
    	avoid divide by 0 when PT = 0

    ks	26. oct. 2008	rev 1.3
    	code optimization

    hm	10. mar. 2009	rev 1.4
    	changed real constants to use dot syntax
    *)
END_FUNCTION_BLOCK

(* ---- GEN_SIN.st ---- *)
FUNCTION_BLOCK GEN_SIN
    (*http://www.oscat.de/images/OSCATBasic/oscat_basic333_en.pdf#page=261*)
    (* read system time and prepare input data *)
    tx := UDINT_TO_TIME(T_PLC_MS()) - last;
    DL := MODR(DL,1.0);
    IF DL < 0.0 THEN DL := 1.0 - DL; END_IF

    (* init section *)
    IF NOT init THEN
    	init := TRUE;
    	last := tx;
    	tx := t#0s;
    END_IF

    (* add last if one cycle is finished *)
    IF tx >= PT THEN
    	last := last + PT;
    	tx := tx - PT;
    END_IF

    (* generate sine wave *)
    IF PT > t#0s THEN temp := SIN(cPI2 * UDINT_TO_REAL(TIME_TO_UDINT(tx + MULTIME(PT, DL))) / UDINT_TO_REAL(TIME_TO_UDINT(PT))); END_IF
    OUT := AM * 0.5 *  temp + OS;

    (* boolean output Q *)
    Q := NOT SIGN_R(temp);

    (* revision history
    hm	22. jan 2007	rev 1.0
    	original version

    hm	17 sep 2007	rev 1.1
    	replaced time() with t_plc_ms for compatibilitx reasons

    hm	27. nov 2007	rev 1.2
    	avoid divide by 0 when PT = 0

    hm	6. jan 2008		rev 1.3
    	improved performance

    hm	16. mar. 2008	rev 1.4
    	added type conversion to avoid warnings under codesys 3.0

    hm	18. oct. 2008	rev 1.5
    	using math constants

    hm	11. mar. 2009	rev 1.6
    	changed real constants to use dot syntax

    *)
END_FUNCTION_BLOCK

(* ---- GEN_SQ.st ---- *)
FUNCTION_BLOCK GEN_SQ
    (*http://www.oscat.de/images/OSCATBasic/oscat_basic333_en.pdf#page=197*)
    (* read system time *)
    tx := T_PLC_MS();

    IF NOT init THEN
    	init := TRUE;
    	tn := tx;
    	Q := TRUE;
    ELSIF tx - tn >= SHR(TIME_TO_UDINT(PT),1) THEN
    	Q := NOT Q;
    	tn := tn + SHR(TIME_TO_UDINT(PT),1);
    END_IF

    (* revision history
    hm	4. aug 2006	rev 1.0
    	original version

    hm	17. sep 2007	rev 1.1
    	replaced time() with T_PLC_MS() for compatibility reasons

    hm	18. jul. 2009	rev 1.2
    	improved accuracy

    hm	16. feb 2011	rev 1.3
    	corrected an error with timer overflow
    *)

END_FUNCTION_BLOCK

(* ---- GEN_SQR.st ---- *)
FUNCTION_BLOCK GEN_SQR
    (*http://www.oscat.de/images/OSCATBasic/oscat_basic333_en.pdf#page=262*)
    (* check DC = 1 or 0 *)
    IF DC = 0.0 THEN
    	OUT := -AM * 0.5 + OS;
    	Q := FALSE;
    	RETURN;
    ELSIF DC = 1.0 THEN
    	OUT := AM * 0.5 + OS;
    	Q := TRUE;
    	RETURN;
    END_IF

    (* read system time and prepare input data *)
    tx := UDINT_TO_TIME(T_PLC_MS()) - last;
    DL := MODR(DL,1.0);
    IF DL < 0.0 THEN DL := 1.0 - DL; END_IF
    DC := MODR(DC,1.0);
    IF DC < 0.0 THEN DC := 1.0 - DC; END_IF

    (* init section *)
    IF NOT init THEN
    	init := TRUE;
    	last := tx;
    	tx := t#0s;
    END_IF

    (* add last if one cycle is finished *)
    IF tx >= PT THEN
    	last := last + PT;
    	tx := tx - PT;
    END_IF

    (* check if falling or rising edge first *)
    IF MULTIME(PT, DL + DC) >= PT THEN
    	(* generate falling edge *)
    	IF tx >= MULTIME(PT, DL + DC - 1) THEN
    		OUT := -AM * 0.5 + OS;
    		Q := FALSE;
    	END_IF
    	(* generate rising edge *)
    	IF tx >= MULTIME(PT, DL) THEN
    		OUT := AM * 0.5 + OS;
    		Q := TRUE;
    	END_IF
    ELSE
    	(* generate rising edge first *)
    	IF tx >= MULTIME(PT, DL) THEN
    		OUT := AM * 0.5 + OS;
    		Q := TRUE;
    	END_IF
    	(* generate falling edge *)
    	IF tx >= MULTIME(PT, DL + DC) THEN
    		OUT := -AM * 0.5 +OS;
    		Q := FALSE;
    	END_IF
    END_IF

    (* revision history

    hm	12. feb 2007	rev 1.1
    	added default value for DC = 0.5

    hm	17 sep 2007	rev 1.2
    	replaced time() with t_plc_ms for compatibilitx reasons

    hm	6. jan 2008	rev 1.3
    	improved performance

    hm	11. mar. 2009	rev 1.4
    	changed real constants to use dot syntax
    	set default amplitude to 1.0

    *)

END_FUNCTION_BLOCK

(* ---- HOLIDAY.st ---- *)
FUNCTION_BLOCK HOLIDAY
    (*http://www.oscat.de/images/OSCATBasic/oscat_basic333_en.pdf#page=123*)
    (* for performance reasons only activate once a day *)
    IF last_active = DATE_IN THEN RETURN; END_IF
    last_active := DATE_IN;

    (* determine language *)
    IF LANGU = 0 THEN
    	lx := cLANGUAGE_DEFAULT;
    ELSE
    	lx := MIN(cLANGUAGE_LMAX, LANGU);
    END_IF

    (* berechnung von ostern für das aktuelle jahr *)
    jahr := YEAR_OF_DATE(DATE_IN);
    ostern := EASTER(jahr);
    wdx := DAY_OF_WEEK(DATE_IN);
    Y := FALSE;

    (* check for HOLIDAYS *)
    FOR i := 0 TO SIZE DO
    	x_date := SET_DATE(jahr, HOLIDAYS[i].MONTH , HOLIDAYS[i].DAY);
    	IF HOLIDAYS[i].USE = 1 AND HOLIDAYS[i].MONTH > 0 THEN
    		(* check for fixed date holiday *)
    		IF x_date = DATE_IN THEN
    			Y := TRUE;
    			NAME := HOLIDAYS[i].NAME;
    			RETURN;
    		END_IF
    	ELSIF HOLIDAYS[i].USE = 1 AND HOLIDAYS[i].MONTH = 0 THEN
    		(* check for holiday in reference to easter *)
    		IF DATE_ADD(ostern, HOLIDAYS[i].DAY ,0,0,0) = DATE_IN THEN
    			Y := TRUE;
    			NAME := HOLIDAYS[i].NAME;
    			RETURN;
    		END_IF
    	ELSIF HOLIDAYS[i].USE < 0 THEN
    		(* check for holiday on a weekday before date *)
    		IF DAY_OF_WEEK(DATE_IN) = ABS(HOLIDAYS[i].USE) AND DATE_IN < x_date AND DATE_IN >= DATE_ADD(x_date,-7,0,0,0) THEN
    			Y := TRUE;
    			NAME := HOLIDAYS[i].NAME;
    			RETURN;
    		END_IF
    	END_IF
    END_FOR

    (* check array if today is weekend *)
    IF NOT Y AND (wdx = 5 AND FRIDAY OR wdx = 6 AND SATURDAY OR wdx = 7 AND SUNDAY) THEN
    	Y := TRUE;
    	NAME := cWEEKDAYS[cLANGUAGE[lx],wdx];
    ELSE
    	NAME := '';
    END_IF

    (*
    Neujahrstag 	1. Januar 	• 	• 	• 	• 	• 	• 	• 	• 	• 	• 	• 	• 	• 	• 	• 	•
    Heilige Drei Könige 	6. Januar 	• 	• 												•
    Karfreitag 	Ostersonntag - 2d 	• 	• 	• 	• 	• 	• 	• 	• 	• 	• 	• 	• 	• 	• 	• 	•
    Ostersonntag 	siehe Osterdatum 				(•)
    Ostermontag 	Ostersonntag + 1d 	• 	• 	• 	• 	• 	• 	• 	• 	• 	• 	• 	• 	• 	• 	• 	•
    Tag der Arbeit 	1. Mai 	• 	• 	• 	• 	• 	• 	• 	• 	• 	• 	• 	• 	• 	• 	• 	•
    Christi Himmelfahrt 	Ostersonntag + 39d 	• 	• 	• 	• 	• 	• 	• 	• 	• 	• 	• 	• 	• 	• 	• 	•
    Pfingstsonntag 	Ostersonntag + 49d 				(•)
    Pfingstmontag 	Ostersonntag + 50d 	• 	• 	• 	• 	• 	• 	• 	• 	• 	• 	• 	• 	• 	• 	• 	•
    Fronleichnam 	Ostersonntag + 60d 	• 	• 					• 			• 	• 	• 	1) 			2)
    Augsburger Friedensfest 	8. August 		(3)
    Mariä Himmelfahrt 	15. August 		(5) 										•
    Tag der Deutschen Einheit 	3. Oktober 6) 	• 	• 	• 	• 	• 	• 	• 	• 	• 	• 	• 	• 	• 	• 	• 	•
    Reformationstag 	31. Oktober 				• 				• 					• 	• 		•
    Allerheiligen 	1. November 	• 	• 								• 	• 	•
    Buß- und Bettag 4) 	Mittwoch vor dem 23.11. 			7 										•
    1. Weihnachtstag 	25. Dezember 	• 	• 	• 	• 	• 	• 	• 	• 	• 	• 	• 	• 	• 	• 	• 	•
    2. Weihnachtstag 	26. Dezember 	• 	• 	• 	• 	• 	• 	• 	• 	• 	• 	• 	• 	• 	• 	• 	•
    *)

    (* revision history
    hm 	27. feb. 2007	rev 1.1
    	deleted unused variable init

    hm	31. oct. 2007	rev 1.2
    	changed holiday definition from constant to input constant to allow easier changes by user without recompilation of the lib

    hm 	24. nov. 2007	rev 1.3
    	changes F_use of  Buß_und_Bettag to 0 because this is no official holiday

    hm	7. apr. 2008	rev 1.4
    	improved performance

    hm	7. oct. 2008	rev 1.5
    	changed code to use setup data from global constants
    	changed length of output NAME from 20 to 30
    	holiday will now also be indicated on a weekend
    	changed function year to year_of_date
    	changed function weekday to day_of_week

    hm	21. oct. 2008	rev 1.6
    	using location constants

    hm	18. jan 2011	rev 2.0
    	using user specified array for HOLIDAYS

    *)

END_FUNCTION_BLOCK

(* ---- HYST.st ---- *)
FUNCTION_BLOCK HYST
    (*http://www.oscat.de/images/OSCATBasic/oscat_basic333_en.pdf#page=421*)
    IF ON >= OFF THEN
    	IF IN < OFF THEN
    		Q := FALSE;
    		WIN := FALSE;
    	ELSIF  IN > ON THEN
    		Q := TRUE;
    		WIN := FALSE;
    	ELSE
    		WIN := TRUE;
    	END_IF
    ELSE
    	IF IN > OFF THEN
    		Q := FALSE;
    		WIN := FALSE;
    	ELSIF  IN < ON THEN
    		Q := TRUE;
    		WIN := FALSE;
    	ELSE
    		WIN := TRUE;
    	END_IF
    END_IF

    (* revision history
    hm		2.  jun 2008	rev 1.0
    	original version

    *)
END_FUNCTION_BLOCK

(* ---- HYST_1.st ---- *)
FUNCTION_BLOCK HYST_1
    (*http://www.oscat.de/images/OSCATBasic/oscat_basic333_en.pdf#page=422*)
    IF IN < LOW THEN
    	Q := FALSE;
    	WIN := FALSE;
    ELSIF IN > HIGH THEN
    	Q := TRUE;
    	WIN := FALSE;
    ELSE
    	WIN := TRUE;
    END_IF

    (* revision history
    hm		4.  aug. 2006	rev 1.0
    	original version

    hm		2. jun. 2008	rev 1.1
    	improved performance
    *)
END_FUNCTION_BLOCK

(* ---- HYST_2.st ---- *)
FUNCTION_BLOCK HYST_2
    (*http://www.oscat.de/images/OSCATBasic/oscat_basic333_en.pdf#page=424*)
    tmp := VAL - HYS * 0.5;
    IF IN < tmp THEN
    	Q := FALSE;
    	WIN := FALSE;
    ELSIF IN > tmp + HYS THEN
    	Q := TRUE;
    	WIN := FALSE;
    ELSE
    	WIN := TRUE;
    END_IF

    (* revision history
    hm		4. aug 2006	rev 1.0
    	original version

    hm		5. jan 2008	rev 1.1
    	improved code for better performance

    hm		2. jun. 2008	rev 1.2
    	improved performance
    *)
END_FUNCTION_BLOCK

(* ---- HYST_3.st ---- *)
FUNCTION_BLOCK HYST_3
    (*http://www.oscat.de/images/OSCATBasic/oscat_basic333_en.pdf#page=425*)
    X := HYST * 0.5;
    IF IN < VAL1 - X THEN
    	Q1 := TRUE;
    ELSIF IN > VAL1 + X THEN
    	Q1 := FALSE;
    END_IF
    IF IN < VAL2 - X THEN
    	Q2 := FALSE;
    ELSIF IN > VAL2 + X THEN
    	Q2 := TRUE;
    END_IF

    (* revision history
    hm	22. jan 2007	rev 1.0
    	original version

    hm	27. dec 2007	rev 1.1
    	changed code for better performance

    hm	5. jan 2008	rev 1.2
    	further performance iprovements

    *)

END_FUNCTION_BLOCK

(* ---- INC_DEC.st ---- *)
FUNCTION_BLOCK INC_DEC
    (*http://www.oscat.de/images/OSCATBasic/oscat_basic333_en.pdf#page=459*)
    axb := CHA XOR CHB;

    (* create pulses for channel a *)
    clka := CHA XOR edgea;
    edgea := CHA;

    clkb := CHB XOR edgeb;
    edgeb := CHB;

    (* create pulses for both channels *)
    clk := clka OR clkb;

    (* set the direction output *)
    IF axb AND clka THEN DIR := TRUE; END_IF
    IF axb AND clkb THEN DIR := FALSE; END_IF

    (* increment or decrement the counter *)
    IF clk AND DIR THEN CNT := CNT + 1; END_IF
    IF clk AND NOT DIR THEN CNT := CNT -1; END_IF

    (* reset the counter if RST active *)
    IF RST THEN CNT := 0; END_IF

END_FUNCTION_BLOCK

(* ---- INTEGRATE.st ---- *)
FUNCTION_BLOCK INTEGRATE
    (*http://www.oscat.de/images/OSCATBasic/oscat_basic333_en.pdf#page=426*)
    (*read system time *)
    tx := T_PLC_MS();

    IF NOT init THEN
    	init := TRUE;
    	X_last := X;
    ELSIF E THEN
    	Y := (X + X_last) * 0.5E-3 * UDINT_TO_REAL(tx-last) * K + Y;
    	X_last := X;
    END_IF
    last := tx;

    (*
    hm 3. nov. 2008	rev 1.0
    original version

    *)

END_FUNCTION_BLOCK

(* ---- INTERLOCK.st ---- *)
FUNCTION_BLOCK INTERLOCK
    (*http://www.oscat.de/images/OSCATBasic/oscat_basic333_en.pdf#page=461*)
    (* the input signal have a run delay to lockout the other input *)
    T1(IN := I1, PT := TL);
    T2(IN := I2, PT := TL);

    Q1 := I1 AND NOT T2.Q;
    Q2 := I2 AND NOT T1.Q;

    (* revision history

    hm	28 sep 2007		rev 1.0
    	original version

    *)
END_FUNCTION_BLOCK

(* ---- INTERLOCK_4.st ---- *)
FUNCTION_BLOCK INTERLOCK_4
    (*http://www.oscat.de/images/OSCATBasic/oscat_basic333_en.pdf#page=462*)
    (* check if enable is active *)
    IF E THEN
    (* reset all vars when there is a MODE change on thy fly *)
    	IF MODE <> lmode THEN
    		OUT := 0;
    		last := 0;
    		old := 0;
    		lmode := MODE;
    	END_IF
    	(* load inputs into in *)
    	in.0 := I0;
    	in.1 := I1;
    	in.2 := I2;
    	in.3 := I3;
    	(* only execute when there is any change *)
    	IF in <> last THEN
    		(* only execute when inputs have chages state *)
    		CASE MODE OF
    			0:	(* output directly display inputs as bits in byte OUT *)
    				OUT := in;

    			1:	(* the input with the highest number will be acepted *)
    				IF in.3 THEN OUT := 8;
    				ELSIF in.2 THEN OUT := 4;
    				ELSIF in.1 THEN OUT := 2;
    				ELSE OUT := in;
    				END_IF

    			2:	(* input last pressed will be displayed only *)
    				last := ((in XOR last) AND in);
    				IF last.3 THEN OUT := 8;
    				ELSIF last.2 THEN OUT := 4;
    				ELSIF last.1 THEN OUT := 2;
    				ELSE OUT := last;
    				END_IF

    			3:	(* any input active will disable all other inputs *)
    				IF (OUT AND in) = 0 THEN
    					IF in.3 THEN OUT := 8;
    					ELSIF in.2 THEN OUT := 4;
    					ELSIF in.1 THEN OUT := 2;
    					ELSE OUT := in;
    					END_IF
    				END_IF

    		END_CASE
    		last := in;
    	END_IF
    	TP := OUT <> old;
    	old := OUT;
    ELSE
    	OUT := 0;
    	last := 0;
    	old := 0;
    	lmode := 0;
    	TP := FALSE;
    END_IF

    (* revision history
    hm	24. oct 2008	rev 1.0
    	original version

    hm	14. mar. 2009	rev 1.1
    	replaced double assignments

    *)
END_FUNCTION_BLOCK

(* ---- LENGTH.st ---- *)
FUNCTION_BLOCK LENGTH
    (*http://www.oscat.de/images/OSCATBasic/oscat_basic333_en.pdf#page=367*)
    YM :=	M
    		+ P * 0.000376065
    		+ IN * 0.0254
    		+ FT * 0.3048
    		+ YD * 0.9144
    		+ MILE * 1609.344
    		+ SM * 1852.0
    		+ FM * 1.829;
    YP := YM * 2659.11478068951;
    YIN := YM * 39.37007874016;
    YFT := YM * 3.28083989501;
    YYD := YM * 1.09361329834;
    YMILE := YM * 0.00062137119;
    YSM := YM * 0.00053995680;
    YFM := YM * 0.54674685621;

    (*
    Länge Meter M SI-Basiseinheit
    Astronomische Einheit* AE 1 AE = 149,597 870 · E9 M
    Parsec pc 1 pc = 206265 AE = 30,857 · E15 M
    Lichtjahr Lj 1 Lj = 9,460 530 · E15 M = 63240 AE = 0,306 59 pc
    Ångström Å 1 Å = E–l0 M
    typograph. Punkt P 1 P = 0,376 065 mm • im Druckereigewerbe
    inch** IN 1 IN = 2,54 · E–2 M = 25,4 mm***
    foot FT 1 FT = 0,3048 M = 30,48 cm
    yard YD 1 YD = 0,9144 M
    MILE MILE 1 MILE = 1609,344 M
    Internat. Seemeile SM 1 SM = 1852 M
    Fathom FM 1 FM = 1,829 M • IN der Seeschifffahrt
    *)

    (* revision history

    hm	27. mar. 2007	rev 1.0
    	original version

    hm	11. mar. 2009	rev 1.1
    	improved code

    *)

END_FUNCTION_BLOCK

(* ---- LIST_NEXT.st ---- *)
FUNCTION_BLOCK LIST_NEXT
    (*http://www.oscat.de/images/OSCATBasic/oscat_basic333_en.pdf#page=487*)
    pt ACCESS ADR(LIST);
    po ACCESS ADR(LEL);

    IF RST THEN
    	pos := 1;
    END_IF

    IF pt[pos] = 0 OR pos = LIST_LENGTH THEN
    	LEL := '';
    	NUL := TRUE;
    ELSE
    	NUL := FALSE;
    	write := 1;
    	FOR pos := pos + 1 TO LIST_LENGTH DO
    		c := pt[pos];
    		IF c = 0 OR c = SEP THEN
    			po[write] := 0;
    			RETURN;
    		ELSE
    			po[write] := pt[pos];
    			write := write + 1;
    		END_IF
    	END_FOR
    END_IF

    (* revision histroy
    hm	25. jun. 2008	rev 1.0
    	original release

    hm	19. jan. 2011	rev 1.1
    	changed string(255) to string(LIST_LENGTH)

    hm	21. mar. 2011	rev 2.0
    	all elements start with SEP

    *)

END_FUNCTION_BLOCK

(* ---- LTCH.st ---- *)
FUNCTION_BLOCK LTCH
    (*http://www.oscat.de/images/OSCATBasic/oscat_basic333_en.pdf#page=242*)
    (* as long as L is true, the latch is transparent and and change of D is transferred to Q *)
    (* of course only when there is no asynchronous reset *)
    IF RST THEN				(* if asynchronous reset then Q=0 *)
    	Q := FALSE;
    ELSIF L THEN			(* latch is transparent *)
    	Q := D;
    END_IF

    (* revision history
    hm	4. aug 2006		rev 1.0
    	original version

    hm	27. dec 2007	rev 1.1
    	changed code for better performance

    hm	30. oct. 2008	rev 1.2
    	deleted unnecessary init with 0

    *)
END_FUNCTION_BLOCK

(* ---- LTCH_4.st ---- *)
FUNCTION_BLOCK LTCH_4
    (*http://www.oscat.de/images/OSCATBasic/oscat_basic333_en.pdf#page=246*)
    (* as long as L is true, the latch is transparent and and change of D is transferred to Q *)
    (* of course only when there is no asynchronous reset *)
    IF RST THEN			(* if asynchronous reset then Q=0 *)
    	Q0 := FALSE;
    	Q1 := FALSE;
    	Q2 := FALSE;
    	Q3 := FALSE;
    ELSIF L THEN			(* latch is transparent *)
    	Q0 := D0;
    	Q1 := D1;
    	Q2 := D2;
    	Q3 := D3;
    END_IF

    (* revision history
    hm	4. aug 2006	rev 1.0
    	original version

    hm	27. dec 2007	rev 1.1
    	changed code for better performance

    hm	30. oct. 2008	rev 1.2
    	deleted unnecessary init with 0

    hm	14. mar. 2009	rev 1.3
    	removed double assignments

    *)
END_FUNCTION_BLOCK

(* ---- M_D.st ---- *)
FUNCTION_BLOCK M_D
    (*http://www.oscat.de/images/OSCATBasic/oscat_basic333_en.pdf#page=341*)
    (* check for RST input *)
    IF RST OR ET >= TMAX THEN
    	PT := t#0ms;
    	ET := t#0ms;
    	startup := FALSE;
    	RUN := FALSE;
    END_IF

    (* avoid timers to START when input is true at startup *)
    IF NOT startup THEN
    	edge_ := START;
    	startup := TRUE;
    END_IF

    (* read system timer *)
    tx := UDINT_TO_TIME(T_PLC_MS());

    (* detect rising edge_ on START *)
    IF START AND NOT edge_ AND NOT STOP THEN
    	T0 := tx;
    	RUN := TRUE;
    	PT := t#0s;
    ELSIF STOP AND RUN THEN
    	PT := ET;
    	RUN := FALSE;
    END_IF
    edge_ := START;
    IF RUN THEN ET := tx - T0; END_IF

    (* revision history
    hm		2.5.2007	rev 1.0
    	original version

    hm		16.9.2007	rev 1.1
    	changes time() to T_plc_ms() for compatibility reasons

    hm	27. feb 2009	rev 1.2
    	deleted unnecessary init with 0
    *)

END_FUNCTION_BLOCK

(* ---- M_T.st ---- *)
FUNCTION_BLOCK M_T
    (*http://www.oscat.de/images/OSCATBasic/oscat_basic333_en.pdf#page=342*)
    (* read system time *)
    tx := UDINT_TO_TIME(T_PLC_MS());

    IF RST OR ET >= TMAX THEN
    	PT :=  t#0s;
    	ET := t#0s;
    ELSIF IN THEN
    	IF NOT edge_ THEN start := tx; END_IF
    	ET := tx - start;
    ELSE
    	PT := ET;
    END_IF
    edge_ := IN;

    (* revision history
    hm	4. aug. 2006	rev 1.0
    	original version

    hm	2. may. 2007	rev 1.1
    	added init variable to avoid unreasonable measurement if falling edge_ occurs first.
    	added ET (elapsed time) output to count from 0 at rising edge_ until a falling edge_ resets ET to 0.
    	added reset input.

    hm	16. sep. 2007	rev 1.2
    	changes time() to T_plc_ms() for compatibility reasons

    hm	17. dec. 2008	rev 1.3
    	code optimized

    hm	10. mar. 2009	rev 1.4
    	removed nested comments
    	removed double assignments

    *)
END_FUNCTION_BLOCK

(* ---- M_TX.st ---- *)
FUNCTION_BLOCK M_TX
    (*http://www.oscat.de/images/OSCATBasic/oscat_basic333_en.pdf#page=342*)
    (* check FOR RST input *)
    IF RST OR (ET >= TMAX) THEN
    	rise := FALSE;
    	fall := FALSE;
    	startup := FALSE;
    	TH := t#0ms;
    	TL := t#0ms;
    	DC := 0.0;
    	F := 0.0;
    	ET := t#0s;
    END_IF

    (* avoid timers to start when input is true at startup *)
    IF NOT startup THEN
    	edge_ := IN;
    	startup := TRUE;
    END_IF

    (* read system timer *)
    tx := UDINT_TO_TIME(T_PLC_MS());

    (* edge_ trigger rising and falling edge_ *)
    IF IN XOR edge_ THEN
    	edge_ := IN;
    	(* rising edge_ starts measurement *)
    	IF IN THEN
    		start := tx;
    		rise := TRUE;
    		IF fall THEN TL := start - stop; END_IF
    		IF TH > t#0ms AND TL > t#0ms THEN
    			DC := TIME_TO_REAL(TH) / TIME_TO_REAL(TH+TL);
    			F := 1000.0 / TIME_TO_REAL(TH + TL);
    		END_IF
    	(* falling edge_ starts second cycle measurement *)
    	ELSE
    		stop := tx;
    		fall := TRUE;
    		IF rise THEN TH := stop - start; END_IF
    		IF TH > t#0ms AND TL > t#0ms THEN
    			DC := TIME_TO_REAL(TH) /  TIME_TO_REAL(TH+TL);
    			F := 1000.0 / TIME_TO_REAL(TH + TL);
    		END_IF
    	END_IF
    END_IF
    IF rise THEN ET := tx - start; END_IF

    (* revision history
    hm	4. aug. 2006	rev 1.0
    	original version

    hm	2. mai. 2007	rev 1.1
    	made sure that no undefined values would be measured at startup conditions
    	added output ET
    	added RST input
    	added TMAX input

    hm	16. sep. 2007	rev 1.2
    	changes time() to T_plc_ms() for compatibility reasons

    hm	27. feb. 2009	rev 1.3
    	deleted unnecessary init with 0

    hm	11. mar. 2009	rev 1.4
    	changed real constants to use dot syntax

    *)
END_FUNCTION_BLOCK

(* ---- MANUAL_1.st ---- *)
FUNCTION_BLOCK MANUAL_1
    (*http://www.oscat.de/images/OSCATBasic/oscat_basic333_en.pdf#page=464*)
    IF NOT MAN THEN
    	Q := IN;
    	STATUS := 100;
    	edge_ := FALSE;
    ELSIF NOT S_edge AND SET THEN
    	Q := TRUE;
    	edge_ := TRUE;
    	STATUS := 101;
    ELSIF NOT r_edge AND RST THEN
    	Q := FALSE;
    	edge_ := TRUE;
    	STATUS := 102;
    ELSIF NOT edge_ THEN
    	Q := M_I;
    	STATUS := 103;
    END_IF

    (* remember levels of manual signals *)
    S_edge := SET;
    r_edge := RST;

    (* revision history
    hm	17. jun 2008	rev 1.0
    	original version

    hm	17. oct 2008	rev 1.1
    	deleted unnecessary variable m_edge

    hm	14. mar. 2009	rev 1.2
    	replaced double assignments

    *)
END_FUNCTION_BLOCK

(* ---- MANUAL_2.st ---- *)
FUNCTION_BLOCK MANUAL_2
    (*http://www.oscat.de/images/OSCATBasic/oscat_basic333_en.pdf#page=464*)
    IF ENA THEN
    	IF NOT ON AND NOT OFF THEN
    		Q := IN;
    		STATUS := 100;
    	ELSIF ON AND NOT OFF THEN
    		Q := TRUE;
    		STATUS := 101;
    	ELSIF NOT ON AND OFF THEN
    		Q := FALSE;
    		STATUS := 102;
    	ELSE
    		Q := MAN;
    		STATUS := 103;
    	END_IF
    ELSE
    	Q := FALSE;
    	STATUS := 104;
    END_IF

    (* revision history
    hm	22. sep. 2008		rev 1.0
    	original version

    *)
END_FUNCTION_BLOCK

(* ---- MANUAL_4.st ---- *)
FUNCTION_BLOCK MANUAL_4
    (*http://www.oscat.de/images/OSCATBasic/oscat_basic333_en.pdf#page=465*)
    IF MAN THEN
    	IF NOT tog THEN
    		Q0 := M0;
    		Q1 := M1;
    		Q2 := M2;
    		Q3 := M3;
    		STATUS := 101;
    	END_IF
    	IF STP AND NOT edge_ THEN
    		tog := TRUE;
    		CASE pos OF
    			0:	Q0 := TRUE;
    				Q1 := FALSE;
    				Q2 := FALSE;
    				Q3 := FALSE;
    				STATUS := 110;
    			1:	Q0 := FALSE;
    				Q1 := TRUE;
    				Q2 := FALSE;
    				Q3 := FALSE;
    				STATUS := 111;
    			2:	Q0 := FALSE;
    				Q1 := FALSE;
    				Q2 := TRUE;
    				Q3 := FALSE;
    				STATUS := 112;
    			3:	Q0 := FALSE;
    				Q1 := FALSE;
    				Q2 := FALSE;
    				Q3 := TRUE;
    				STATUS := 113;
    		END_CASE
    		pos := INC(pos,1,3);
    	END_IF
    ELSE
    	Q0 := I0;
    	Q1 := I1;
    	Q2 := I2;
    	Q3 := I3;
    	STATUS := 100;
    	tog := FALSE;
    	pos := 0;
    END_IF

    (* remember STATUS of STP *)
    edge_ := STP;

    (* revision history
    hm	17. jun 2008		rev 1.0
    	original version

    *)
END_FUNCTION_BLOCK

(* ---- MATRIX.st ---- *)
FUNCTION_BLOCK MATRIX
    (*http://www.oscat.de/images/OSCATBasic/oscat_basic333_en.pdf#page=227*)
    TP := FALSE;
    CODE := 0;
    (* read scan lines *)
    X[line].0 := X1;
    X[line].1 := X2;
    X[line].2 := X3;
    X[line].3 := X4;
    X[line].4 := X5;

    (* compare for change *)
    FOR i := 0 TO 3 DO
    	IF X[i] <> L[i] THEN
    		(* scan line information has changed CODE need to be found and generated *)
    		temp := X[i] XOR L[i];
    		IF temp.0 THEN
    			CODE := 1;
    			CODE.7 := X[i].0;
    			L[i].0 := X[i].0;
    		ELSIF temp.1 THEN
    			CODE := 2;
    			CODE.7 := X[i].1;
    			L[i].1 := X[i].1;
    		ELSIF temp.2 THEN
    			CODE := 3;
    			CODE.7 := X[i].2;
    			L[i].2 := X[i].2;
    		ELSIF temp.3 THEN
    			CODE := 4;
    			CODE.7 := X[i].3;
    			L[i].3 := X[i].3;
    		ELSIF temp.4 THEN
    			CODE := 5;
    			CODE.7 := X[i].4;
    			L[i].4 := X[i].4;
    		END_IF
    		TP := TRUE;
    		CODE.4 := line.0;
    		CODE.5 := line.1;
    		CODE.6 := line.2;

    		(* check if RELEASE codes need to be killed *)
    		IF NOT RELEASE AND CODE < 127 THEN
    			CODE := 0;
    			TP := FALSE;
    		END_IF
    		EXIT;
    	END_IF
    END_FOR

    (* increment scan line every cycle *)
    line := (line + 1) AND 2#0000_0011;
    temp := SHL(BYTE#1,line);
    Y1 := temp.0;
    Y2 := temp.1;
    Y3 := temp.2;
    Y4 := temp.3;

    (* revision history
    hm		10.6.2007	rev 1.0
    	original version

    hm		11.9.2007	rev 1.1
    	deleted unused variables k and old_code

    hm		23.12.2007	rev 1.2
    	added exit statement in for loop instead of i:=5

    hm		26. oct. 2008	rev 1.3
    	CODE optimized

    *)

END_FUNCTION_BLOCK

(* ---- MESSAGE_4R.st ---- *)
FUNCTION_BLOCK MESSAGE_4R
    (*http://www.oscat.de/images/OSCATBasic/oscat_basic333_en.pdf#page=173*)
    (* check for rising edge_ on EN *)
    TR := FALSE;
    IF ENQ THEN
    	IF (NOT edge_ AND CLK) OR timer.Q THEN
    			MN := INC1(MN, MM);
    			TR := TRUE;
    			timer(IN := FALSE);
    			CASE MN OF
    				0 : MX := M0;
    				1 : MX := M1;
    				2 : MX := M2;
    				3 : MX := M3;
    			END_CASE
    	END_IF
    	edge_ := CLK;
    	timer( IN := CLK, PT := T1);
    ELSE
    	MX := '';
    	MN := 0;
    END_IF

    (* revision history
    hm	8. oct. 2008	rev 1.0
    	original version

    hm	27. oct. 2008	rev 1.1
    	changed _INC to INC1

    *)

END_FUNCTION_BLOCK

(* ---- MESSAGE_8.st ---- *)
FUNCTION_BLOCK MESSAGE_8
    (*http://www.oscat.de/images/OSCATBasic/oscat_basic333_en.pdf#page=173*)
    (* check if an alarm is present if yes set the output M otherwise clear M *)
    IF IN1 THEN
    	M := S1;
    ELSIF IN2 THEN
    	M := S2;
    ELSIF IN3 THEN
    	M := S3;
    ELSIF IN4 THEN
    	M := S4;
    ELSIF IN5 THEN
    	M := S5;
    ELSIF IN6 THEN
    	M := S6;
    ELSIF IN7 THEN
    	M := S7;
    ELSIF IN8 THEN
    	M := S8;
    ELSE
    	M := '';
    END_IF

    (* revision history
    hm	26.12.2007		rev 1.0
    	original version

    hm	29. mar. 2008	rev 1.1
    	changed STRING to STRING(STRING_LENGTH)
    *)

END_FUNCTION_BLOCK

(* ---- METER.st ---- *)
FUNCTION_BLOCK METER
    (*http://www.oscat.de/images/OSCATBasic/oscat_basic333_en.pdf#page=343*)
    (* measure the last cycle time and make sure we onle execute once every millisecond *)
    tx := T_PLC_MS();
    IF NOT init THEN
    	init := TRUE;
    	last := tx;
    	MR.RX := MX;
    	MR.R1 := 0.0;
    ELSIF tx = last THEN
    	RETURN;
    ELSE
    	tc := UDINT_TO_REAL(tx - last) * 0.001;
    END_IF
    last := tx;

    (* reset *)
    IF RST THEN
    	MR.R1 := 0.0;
    	MR.RX := 0.0;
    ELSE
    	(* current consumption measurement *)
    	IF I1 THEN MX1 := M1; ELSE MX1 := 0.0; END_IF
    	IF I2 THEN MX2 := M2; ELSE MX2 := 0.0; END_IF
    	(* add up the current values in a double real *)
    	R2_ADD(MR,(SEL(I1,0.0,MX1) + SEL(I2, 0.0, MX2)) / D * tc, MR);
    	(* set the current output value *)
    	MX := MR.RX;
    END_IF

    (* revision history

    hm	16. sep.2007		rev 1.0
    	original version

    hm	7. feb 2008		rev 1.1
    	use new version of ft_int to avoid a counting stop at high values
    	deleted unnecessary limits

    hm	24. mar. 2008	rev 1.2
    	use data_type real2 to extend accuracy to 15 digits total
    	do not use ft_int which adds unnecessary overhead

    hm	8. feb. 2009	rev 1.3
    	changed MX to be I/O
    	make sure calculation works for cycle times < 1 ms

    hm	8. mar. 2009	rev 1.4
    	last was not updated
    	code improvements

    *)

END_FUNCTION_BLOCK

(* ---- METER_STAT.st ---- *)
FUNCTION_BLOCK METER_STAT
    (*http://www.oscat.de/images/OSCATBasic/oscat_basic333_en.pdf#page=345*)
    IF RST THEN
    	LAST_DAY := 0.0;
    	CURRENT_DAY := 0.0;
    	Day_Start := IN;
    	LAST_WEEK := 0.0;
    	CURRENT_WEEK := 0.0;
    	Week_Start := IN;
    	LAST_MONTH := 0.0;
    	CURRENT_MONTH := 0.0;
    	Month_Start := IN;
    	LAST_YEAR := 0.0;
    	CURRENT_YEAR := 0.0;
    	Year_Start := IN;
    ELSE
    	CURRENT_DAY := IN - Day_Start;
    	CURRENT_WEEK := IN - Week_Start;
    	CURRENT_MONTH := IN - Month_Start;
    	CURRENT_YEAR := IN - Year_Start;
    END_IF

    IF YEAR_OF_DATE(DI) > YEAR_OF_DATE(last_run) THEN
    	(* a new year has started *)
    	LAST_YEAR := CURRENT_YEAR;
    	CURRENT_YEAR := 0.0;
    	Year_Start := IN;
    	LAST_MONTH := CURRENT_MONTH;
    	CURRENT_MONTH := 0.0;
    	Month_Start := IN;
    	LAST_DAY := CURRENT_DAY;
    	CURRENT_DAY := 0.0;
    	Day_Start := IN;
    ELSIF MONTH_OF_DATE(DI) > MONTH_OF_DATE(last_run) THEN
    	(* a new month has started, january is alrerady done by year change *)
    	LAST_MONTH := CURRENT_MONTH;
    	CURRENT_MONTH := 0.0;
    	Month_Start := IN;
    	LAST_DAY := CURRENT_DAY;
    	CURRENT_DAY := 0.0;
    	Day_Start := IN;
    ELSIF DAY_OF_YEAR(DI) > DAY_OF_YEAR(last_run) THEN
    	(* day has chaged, first day of year and first day of month has already been taken care of *)
    	LAST_DAY := CURRENT_DAY;
    	CURRENT_DAY := 0.0;
    	Day_Start := IN;
    END_IF
    IF DAY_OF_WEEK(DI) < DAY_OF_WEEK(last_run) THEN
    	(* a new week has started *)
    	LAST_WEEK := CURRENT_WEEK;
    	CURRENT_WEEK := 0.0;
    	Week_Start := IN;
    END_IF
    last_run := DI;

    (* revision history
    hm	16. sep. 2007	rev 1.0
    	original version

    hm	7. oct. 2008	rev 1.1
    	changed function year_to_year_of_date
    	changed function month to month_of_date
    	changed function weekday to day_of_week

    hm	11. mar. 2009	rev 1.2
    	changed real constants to use dot syntax

    hm	18. jul. 2009	rev 1.3
    	changes all outputs to be I/O
    *)

END_FUNCTION_BLOCK

(* ---- ONTIME.st ---- *)
FUNCTION_BLOCK ONTIME
    (*http://www.oscat.de/images/OSCATBasic/oscat_basic333_en.pdf#page=346*)
    (* read system time *)
    tx := T_PLC_MS();

    (* make sure the first cycle works correctly *)
    IF NOT init THEN
    	init := TRUE;
    	last := tx;
    	ms := 0;
    END_IF
    IF RST THEN
    	SECONDS := 0;
    	CYCLES := 0;
    	last := tx;
    	ms := 0;
    ELSIF IN THEN
    	(* add the current milliseconds *)
    	ms := (tx - last) + ms;
    	IF ms >= 1000 THEN
    		SECONDS := SECONDS + 1;
    		ms := ms - 1000;
    	END_IF
    	CYCLES := CYCLES + BOOL_TO_UINT(NOT edge_);
    END_IF
    last := tx;
    edge_ := IN;

    (* revision history
    hm 22.2.2007		rev 1.1
    	changed VAR RETAIN PERSISTENT to VAR RETAIN for better compatibility
    	wago lon contollers do not support persisitent

    hm 2.8.2007		rev 1.2
    	adding time up IN a real number will automatically lead to the point where
    	small time scales like the cycle time will be below the resolution of real and therefore
    	ontime would not increase IN small steps as necessary
    	the time is now measured internally IN two  UDINTs and be converted to real only for
    	output purposes.
    	deleted the variable power because it was unnecessary

    hm	16.9.2007		rev 1.3
    	changes time() to T_plc_ms() for compatibility reasons

    hm	2. dec. 2007	rev 1.4
    	chaged code for better performance

    hm	16. mar. 2008	rev 1.5
    	added type conversions to avoid warnings under codesys 3.0

    hm	21. oct. 2008	rev 2.0
    	changed module for much better performance and allow for external result storage

    hm	10. nov. 2008	rev 2.1
    	increased internal resolution to milliseconds

    hm	16. nov. 2008	rev 2.2
    	changed typecast to avoid warnings

    hm	17. dec. 2008	rev 2.3
    	fixed an error when IN would be true for more then 49 days

    hm	17. jan 2011	rev 2.4
    	init will not clear SECONDS and CYCLES, only RST clears these values

    hm	18. mar. 2011	rev 2.5
    	reset was not working

    *)
END_FUNCTION_BLOCK
